(* IEC 61131-3 sources: kns-pump-station/tests/POUs/Model/FB_TankModel_Test, 13 files *)

(* ---- FB_TankModel_Test.decl.st ---- *)
// Назначение: набор coUnit для FB_TankModel — баланс объёма резервуара: интегрирование притока и откачки,
//             перелив и его время, осушенный приёмок, шаг 0 и «время назад», установка уровня. Ожидаемые значения —
//             эталон tools_project/plant_reference.py (сценарии tank.*): dh = (Qin − Qout)·dt / 3600 / S.
// Автор:      kr0nsch
// Версия:     0.1.0
// Документ:   docs/DESIGN.md, разделы 11.3, 14.1
FUNCTION_BLOCK FB_TankModel_Test EXTENDS coUnit.FB_TestSuite
VAR CONSTANT
    R_AREA_M2 : REAL := 12.0;
    R_OVERFLOW_M : REAL := 4.6;
    LR_STEP_S : LREAL := 10.0;        // шаг интегрирования в тесте
    LR_SHORT_S : LREAL := 0.2;        // шаг SIM_DT_SUBSTEP
    UI_STEPS_1H : UINT := 360;        // 1 ч шагами по 10 с
    UI_STEPS_10MIN : UINT := 60;
    R_EPS_M : REAL := 1.0E-5;
END_VAR

(* ---- DefaultsLevelAfterSetLevel.method.decl.st ---- *)
// Новый резервуар пуст (уровень 0, приёмок осушен); SetLevel(1,2) и вызов с шагом 0 — уровень 1,2 м,
// объём 14,4 м³, перелива нет.
METHOD PRIVATE DefaultsLevelAfterSetLevel
VAR
    fbDut : FB_TankModel;
END_VAR

(* ---- IntakeDryNoFlow.method.decl.st ---- *)
// Уровень 0,25 м ниже приёмка 0,30 м: откачка 150 м³/ч не уменьшает уровень (насосы подсасывают
// воздух); приток 12 м³/ч 10 мин поднимает уровень на 0,1667 м — приёмок снова под водой.
METHOD PRIVATE IntakeDryNoFlow
VAR
    fbDut : FB_TankModel;       // проверяемый ФБ
    uiI : UINT;
END_VAR

(* ---- IntakeDryNoFlow.method.impl.st ---- *)
coUnit.TEST('TankModel_IntakeDryNoFlow');

fbDut.SetLevel(rNewLevel_m := 0.25);
fbDut(rInflow_m3h := 0.0, rOutflow_m3h := 150.0, lrDt_s := LR_STEP_S, rArea_m2 := R_AREA_M2,
      rOverflow_m := R_OVERFLOW_M);
AssertTrue(Condition := fbDut.xIntakeDry, Message := 'intake dry');
AssertEquals_REAL(Expected := 0.25, Actual := fbDut.rLevel_m, Delta := R_EPS_M, Message := 'no pumping below intake');
FOR uiI := 1 TO UI_STEPS_10MIN DO
    fbDut(rInflow_m3h := 12.0, rOutflow_m3h := 0.0, lrDt_s := LR_STEP_S, rArea_m2 := R_AREA_M2,
          rOverflow_m := R_OVERFLOW_M);
END_FOR
AssertEquals_REAL(Expected := 0.416667, Actual := fbDut.rLevel_m, Delta := R_EPS_M, Message := 'inflow raises level');
AssertFalse(Condition := fbDut.xIntakeDry, Message := 'intake under water again');

coUnit.TEST_FINISHED();

(* ---- NoOverflowWhenBalanced.method.decl.st ---- *)
// На отметке перелива при притоке, равном откачке (150 м³/ч), вода не переливается: уровень 4,6 м держится,
// время перелива не растёт — перелив считается, только пока приток больше откачки.
METHOD PRIVATE NoOverflowWhenBalanced
VAR
    fbDut : FB_TankModel;       // проверяемый ФБ
    uiI : UINT;
END_VAR

(* ---- NoOverflowWhenBalanced.method.impl.st ---- *)
coUnit.TEST('TankModel_NoOverflowWhenBalanced');

fbDut.SetLevel(rNewLevel_m := R_OVERFLOW_M);
FOR uiI := 1 TO 6 DO
    fbDut(rInflow_m3h := 150.0, rOutflow_m3h := 150.0, lrDt_s := LR_STEP_S, rArea_m2 := R_AREA_M2,
          rOverflow_m := R_OVERFLOW_M);
END_FOR
AssertEquals_REAL(Expected := R_OVERFLOW_M, Actual := fbDut.rLevel_m, Delta := R_EPS_M,
                  Message := 'level kept at mark');
AssertFalse(Condition := fbDut.xOverflow, Message := 'no overflow when balanced');
AssertEquals_UDINT(Expected := 0, Actual := fbDut.udiOverflow_s, Message := 'no overflow time');

coUnit.TEST_FINISHED();

(* ---- OverflowCounts.method.decl.st ---- *)
// От 4,5 м при притоке 250 м³/ч без откачки: 0,1 м набирается за 17,3 с, дальше уровень ограничен
// 4,6 м, время перелива растёт по шагам, где приток больше откачки: 59 шагов по 10 с = 590 с.
METHOD PRIVATE OverflowCounts
VAR
    fbDut : FB_TankModel;       // проверяемый ФБ
    uiI : UINT;
END_VAR

(* ---- OverflowCounts.method.impl.st ---- *)
coUnit.TEST('TankModel_OverflowCounts');

fbDut.SetLevel(rNewLevel_m := 4.5);
FOR uiI := 1 TO UI_STEPS_10MIN DO
    fbDut(rInflow_m3h := 250.0, rOutflow_m3h := 0.0, lrDt_s := LR_STEP_S, rArea_m2 := R_AREA_M2,
          rOverflow_m := R_OVERFLOW_M);
END_FOR
AssertEquals_REAL(Expected := R_OVERFLOW_M, Actual := fbDut.rLevel_m, Delta := R_EPS_M,
                  Message := 'level limited at overflow');
AssertTrue(Condition := fbDut.xOverflow, Message := 'overflow active');
AssertEquals_UDINT(Expected := 590, Actual := fbDut.udiOverflow_s, Message := 'overflow seconds');
fbDut(rInflow_m3h := 100.0, rOutflow_m3h := 150.0, lrDt_s := LR_STEP_S, rArea_m2 := R_AREA_M2,
      rOverflow_m := R_OVERFLOW_M);
AssertFalse(Condition := fbDut.xOverflow, Message := 'overflow stops when pumps exceed inflow');
AssertTrue(Condition := fbDut.rLevel_m < R_OVERFLOW_M, Message := 'level falls');
AssertEquals_UDINT(Expected := 590, Actual := fbDut.udiOverflow_s, Message := 'overflow seconds kept');

coUnit.TEST_FINISHED();

(* ---- SetLevelClamped.method.decl.st ---- *)
// SetLevel ограничивает уровень 0…отметка перелива; неконечное значение не принимается.
METHOD PRIVATE SetLevelClamped
VAR
    fbDut : FB_TankModel;       // проверяемый ФБ
    uBits : PL.U_RealBits;
END_VAR

(* ---- ShortOverflowCounted.method.decl.st ---- *)
// Перелив короче 1 с (один шаг 0,2 с на отметке перелива) виден в udiOverflow_s: не меньше 1 с. Иначе
// округление до целых секунд давало бы 0, и проверка «перелива нет (udiOverflow_s = 0)» PMI-20 и PMI-24
// проходила бы при настоящем переливе.
METHOD PRIVATE ShortOverflowCounted
VAR
    fbDut : FB_TankModel;       // проверяемый ФБ
END_VAR

(* ---- VolumeBalance.method.decl.st ---- *)
// Приток 30, откачка 10 м³/ч в течение 1 ч: уровень 1,2 + 20/12 = 2,866667 м.
METHOD PRIVATE VolumeBalance
VAR
    fbDut : FB_TankModel;       // проверяемый ФБ
    uiI : UINT;
END_VAR

(* ---- VolumeBalance.method.impl.st ---- *)
coUnit.TEST('TankModel_VolumeBalance');

fbDut.SetLevel(rNewLevel_m := 1.2);
FOR uiI := 1 TO UI_STEPS_1H DO
    fbDut(rInflow_m3h := 30.0, rOutflow_m3h := 10.0, lrDt_s := LR_STEP_S, rArea_m2 := R_AREA_M2,
          rOverflow_m := R_OVERFLOW_M);
END_FOR
// ref: tank.balance_30_10_1h.level_m
AssertEquals_REAL(Expected := 2.866667, Actual := fbDut.rLevel_m, Delta := R_EPS_M, Message := 'level after 1 h');
AssertEquals_UDINT(Expected := 0, Actual := fbDut.udiOverflow_s, Message := 'no overflow');

coUnit.TEST_FINISHED();

(* ---- ZeroOrNegativeStepNoChange.method.decl.st ---- *)
// Шаг 0 и отрицательный шаг («время назад») не меняют уровень и время перелива.
METHOD PRIVATE ZeroOrNegativeStepNoChange
VAR
    fbDut : FB_TankModel;       // проверяемый ФБ
END_VAR
